// TIA Portal V20 export
// export: Created 2026-10-11T05:25:32.2887143Z, ExportSetting WithDefaults, DisplayName Totally Integrated Automation Portal, DisplayVersion V20, DisplayName TIA Portal Openness, DisplayVersion V20, DisplayName TIA Portal Teamcenter Gateway, DisplayVersion V20, DisplayName TIA Portal Version Control Interface, DisplayVersion V20, DisplayName SINAMICS Startdrive Advanced, DisplayVersion V20 SP1 Update 2, DisplayName SINAMICS Startdrive G110M, G120, G120C, G120D, G120P, G115D, DisplayVersion V20 SP1 Update 2, DisplayName SINAMICS Startdrive G130, G150, S120, S150, SINAMICS MV, G220, S200, S210, DisplayVersion V20 SP1 Update 2, DisplayName STEP 7 Professional, DisplayVersion V20, DisplayName STEP 7 Safety, DisplayVersion V20, DisplayName WinCC Basic/Comfort/Advanced, DisplayVersion V20, DisplayName WinCC Professional, DisplayVersion V20, DisplayName WinCC Unified, DisplayVersion V20
DATA_BLOCK "StationB"   // DB12
VERSION : 0.1
// stored: AutoNumber true, DBAccessibleFromOPCUA true, DBAccessibleFromWebserver true, InstanceOfName FB_DeclarationUnit, InstanceOfType FB
"FB_DeclarationUnit"
   // VAR_INPUT
   //    Execute { ExternalWritable := 'False'} : Bool;
   //    Abort { ExternalWritable := 'False'} : Bool;
   //    Command { ExternalWritable := 'False'} : DInt;
   //    ParCfg { ExternalWritable := 'False'} : "ST_DeclarationParCfg";
   //    ParCmd { ExternalWritable := 'False'} : "ST_DeclarationParCmd";
   //    ParentIndex { ExternalAccessible := 'False'; ExternalVisible := 'False'; ExternalWritable := 'False'} : DInt;
   //    Startup { ExternalAccessible := 'False'; ExternalVisible := 'False'; ExternalWritable := 'False'} : Bool;
   // END_VAR
   // VAR_OUTPUT
   //    Busy { ExternalWritable := 'False'} : Bool;
   //    Done { ExternalWritable := 'False'} : Bool;
   //    Error { ExternalWritable := 'False'} : Bool;
   //    Aborted { ExternalWritable := 'False'} : Bool;
   //    Held { ExternalWritable := 'False'} : Bool;
   //    ErrorID { ExternalWritable := 'False'} : DWord;
   //    Timing { ExternalWritable := 'False'} : "ST_ModuleTiming";
   //    OutCmd { ExternalWritable := 'False'} : "ST_DeclarationOutCmd";
   //    OutImm { ExternalWritable := 'False'} : "ST_UnitProbeImm";
   // END_VAR
   // VAR_IN_OUT
   //    Hal : "ST_DeclarationUnitHal";
   // END_VAR
   // VAR
   //    Status { ExternalWritable := 'False'; S7_SetPoint := 'True'} : "ST_ModuleStatus";
   //    Core { ExternalAccessible := 'False'; ExternalVisible := 'False'; ExternalWritable := 'False'; S7_SetPoint := 'True'} : "FRK_Core";
   //    LatchedParCmd { ExternalAccessible := 'False'; ExternalVisible := 'False'; ExternalWritable := 'False'; S7_SetPoint := 'True'} : "ST_DeclarationParCmd";
   //    Device { ExternalAccessible := 'False'; ExternalVisible := 'False'; ExternalWritable := 'False'; S7_SetPoint := 'True'} : "ST_UnitProbeDevice";
   //    Unit { ExternalAccessible := 'False'; ExternalVisible := 'False'; ExternalWritable := 'False'; S7_SetPoint := 'True'} : "FRK_Unit";
   //    HmiRequest { S7_SetPoint := 'True'} : "ST_HmiRequest";
   //    ModePolicy { ExternalAccessible := 'False'; ExternalVisible := 'False'; ExternalWritable := 'False'; S7_SetPoint := 'True'} : Array[0..6] of "ST_ModePolicy";
   //    Access { ExternalWritable := 'False'; S7_SetPoint := 'True'} : "FRK_Access";
   //    HmiResponse { ExternalWritable := 'False'; S7_SetPoint := 'True'} : "ST_HmiResponse";
   //    ConfigRev { ExternalWritable := 'False'} : UDInt;
   //    ConfigCursor { ExternalAccessible := 'False'; ExternalVisible := 'False'; ExternalWritable := 'False'; S7_SetPoint := 'True'} : "FRK_ConfigCursor";
   //    Part { ExternalWritable := 'False'; S7_SetPoint := 'True'} : "ST_PartContext";
   //    History { ExternalWritable := 'False'; S7_SetPoint := 'True'} : Array[1..16] of "ST_Diagnostic";
   //    HistoryHead { ExternalWritable := 'False'} : Int;
   //    ModeActivePublished { ExternalWritable := 'False'} : DInt;
   //    RunningPublished { ExternalWritable := 'False'} : Bool;
   //    StopPendingPublished { ExternalWritable := 'False'} : Bool;
   //    SupportedModesPublished { ExternalWritable := 'False'} : Array[0..6] of Bool;
   //    GoodCount { ExternalWritable := 'False'} : UDInt;
   //    NokCount { ExternalWritable := 'False'} : UDInt;
   //    ReworkCount { ExternalWritable := 'False'} : UDInt;
   //    NokReason { ExternalWritable := 'False'} : DInt;
   //    Cell { ExternalWritable := 'False'; S7_SetPoint := 'True'} : "FB_DeclarationCell";
   //    Satellite { ExternalWritable := 'False'; S7_SetPoint := 'True'} : "FB_SatelliteUnit";
   // END_VAR
BEGIN
END_DATA_BLOCK
